// TIA Portal project "State Machine Triple-liquid mixing+HMI final version" (V17)

(* hardware
DEVICE "S7-300/ET200M station_1"  S7-300 station
   slot 0: "Rail_0"  Rail  6ES7 390-1***0-0AA0
   slot 2: "PLC_1"  CPU 317-2 PN/DP  6ES7 317-2EK14-0AB0  V3.2
      slot 2: "PROFINET interface_1"  PN-IO
         slot 1: "Port_1"  Port
         slot 2: "Port_2"  Port
   slot 4: "DI 16x24VDC_1"  DI16 x 24VDC  6ES7 321-1BH02-0AA0
   slot 5: "DO 8x24VDC/0.5A_1"  DO8 x 24VDC / 0.5A  6ES7 322-8BF00-0AB0
   slot 6: "AI 4x0/4mA/20mA, Ex_1"  AI4 x 0/4 to 20mA, Ex  6ES7 331-7RD00-0AB0
DEVICE "HMI_1"  TP1200 Comfort Portrait SIPLUS
   slot 0: "HMI_1"  TP1200 Comfort Portrait SIPLUS  6AG1 124-0MC01-4AX0  17.0.0.0
   slot 1: "HMI_RT_1"  TP1200 Comfort Portrait SIPLUS  6AG1 124-0MC01-4AX0  17.0.0.0
   slot 5: "HMI_1.IE_CP_1"  PROFINET Interface  17.0.0.0
      slot 1: "PROFINET Interface_1"  PROFINET Interface
         slot 1: "Port_1"  Port
         slot 2: "Port_2"  Port
   slot 7: "HMI_1.MPI/DP_CP_1"  MPI/DP Interface  17.0.0.0
*)

// ===== PLC "PLC_1"  CPU 317-2 PN/DP =====

VAR_GLOBAL   // PLC tag table "Default tag table"
   "E_stop" AT %I0.0 : Bool;
   "Actual_level" AT %MD0 : Real;
   "RESET_1" AT %I0.1 : Bool;
   "Start_mixing" AT %I0.2 : Bool;
   "Alarm_light" AT %Q0.0 : Bool;
   "Valve_A" AT %Q4.0 : Bool;
   "Valve_B" AT %Q4.1 : Bool;
   "Valve_C" AT %Q4.2 : Bool;
   "Agitator_Q" AT %Q4.3 : Bool;
   "Drain_valve" AT %Q4.4 : Bool;
   "REC_A" AT %MD4 : Real;
   "REC_B" AT %MD8 : Real;
   "REC_C" AT %MD12 : Real;
   "start_empty" AT %I0.3 : Bool;
   "Eroor_code" AT %MW16 : Int;
   "Start_timer" AT %T0 : Timer;
   "start_empty_Timer" AT %T1 : Timer;
   "Reset_timer" AT %T2 : Timer;
   "RAW_Level_sensor" AT %IW288 : Int;
   "Start_batch" AT %M10.1 : Bool;
   "Reset_HMI" AT %M10.2 : Bool;
   "Start-EMpty" AT %M10.3 : Bool;
   "Status" AT %MW20 : Int;
   "Min_level" AT %MD48 : Real;
   "Max_lvl" AT %MD24 : Real;
   "drain_time_WD" AT %MD28 : Time;
   "Agitator_time_WD" AT %MD32 : Time;
   "FIlling_time_WD" AT %MD36 : Time;
   "Agitating_time" AT %MD40 : Time;
   "Batch_done_confirmation" AT %M44.0 : Bool;
   "Rec_approved" AT %M44.1 : Bool;
   "Tank1_active" AT %M18.0 : Bool;
   "Alarm_HMI" AT %M18.1 : Bool;
   "Valv_A_HMI" AT %M18.2 : Bool;
   "Valv_B_HMI" AT %M18.3 : Bool;
   "Valv_C_HMI" AT %M18.4 : Bool;
   "Agit_HMI" AT %M18.5 : Bool;
   "Drain_valv_HMI" AT %M18.6 : Bool;
END_VAR

DATA_BLOCK "batch_variable"   // DB9
{ S7_Optimized_Access := 'FALSE' }
VERSION : 0.1
   VAR
      reciepe_A : Real;
      reciepe_B : Real;
      reciepe_C : Real;
   END_VAR
BEGIN
END_DATA_BLOCK

DATA_BLOCK "Stat machine_DB"   // DB10
{ S7_Optimized_Access := 'FALSE' }
VERSION : 0.1
// stored: InstanceOfName Stat machine
"Stat machine"
BEGIN
END_DATA_BLOCK

FUNCTION_BLOCK "Stat machine"   // FB1, LAD
{ S7_Optimized_Access := 'FALSE' }
VERSION : 0.1
   VAR_INPUT
      "E-Stop" : Bool;
      Actual_level : Real;
      RESET_Cmd : Bool;
      start_mixing : Bool;
      Reciepes_A : Real;
      Reciepes_c : Real;
      Reciepes_B : Real;
      start_empty : Bool;
      wtachDog_time_Drain : Time;
      wtachDog_time_Agitator : Time;
      wtachDog_time_valve : Time;
      Min_level : Real;
      Agitating_time : Time;
      batch_done_confirmation : Bool;
   END_VAR
   VAR_OUTPUT
      Alram_red_light : Bool;
      q_valve_A : Bool;
      q_valve_B : Bool;
      q_valve_C : Bool;
      Agitaor : Bool;
      drain_valve : Bool;
      Error_code : Int;
      Alarm_active : Bool;
      Valve_A_active : Bool;
      Valve_B_active : Bool;
      Valve_C_active : Bool;
      Agitator_active : Bool;
      Drain_valve_active : Bool;
   END_VAR
   VAR_IN_OUT
      iStep_number : Int;
      max_lvl : Real;
      Recrp_approved : Bool;
   END_VAR
   VAR
      Agitator_runnig : Bool;
      Target_1 : Real;
      Target_2 : Real;
      Reset_alrm : Bool;
      Batch_done : Bool;
      "1%_tank_apacity" : Real;
      max_recepes_valuem : Real;
      "15%_Tank_capacity" : Real;
   END_VAR
   VAR_TEMP   // added for the SCL form of the ladder/FBD networks
      _w1 : Bool;
   END_VAR
BEGIN

REGION Network 1
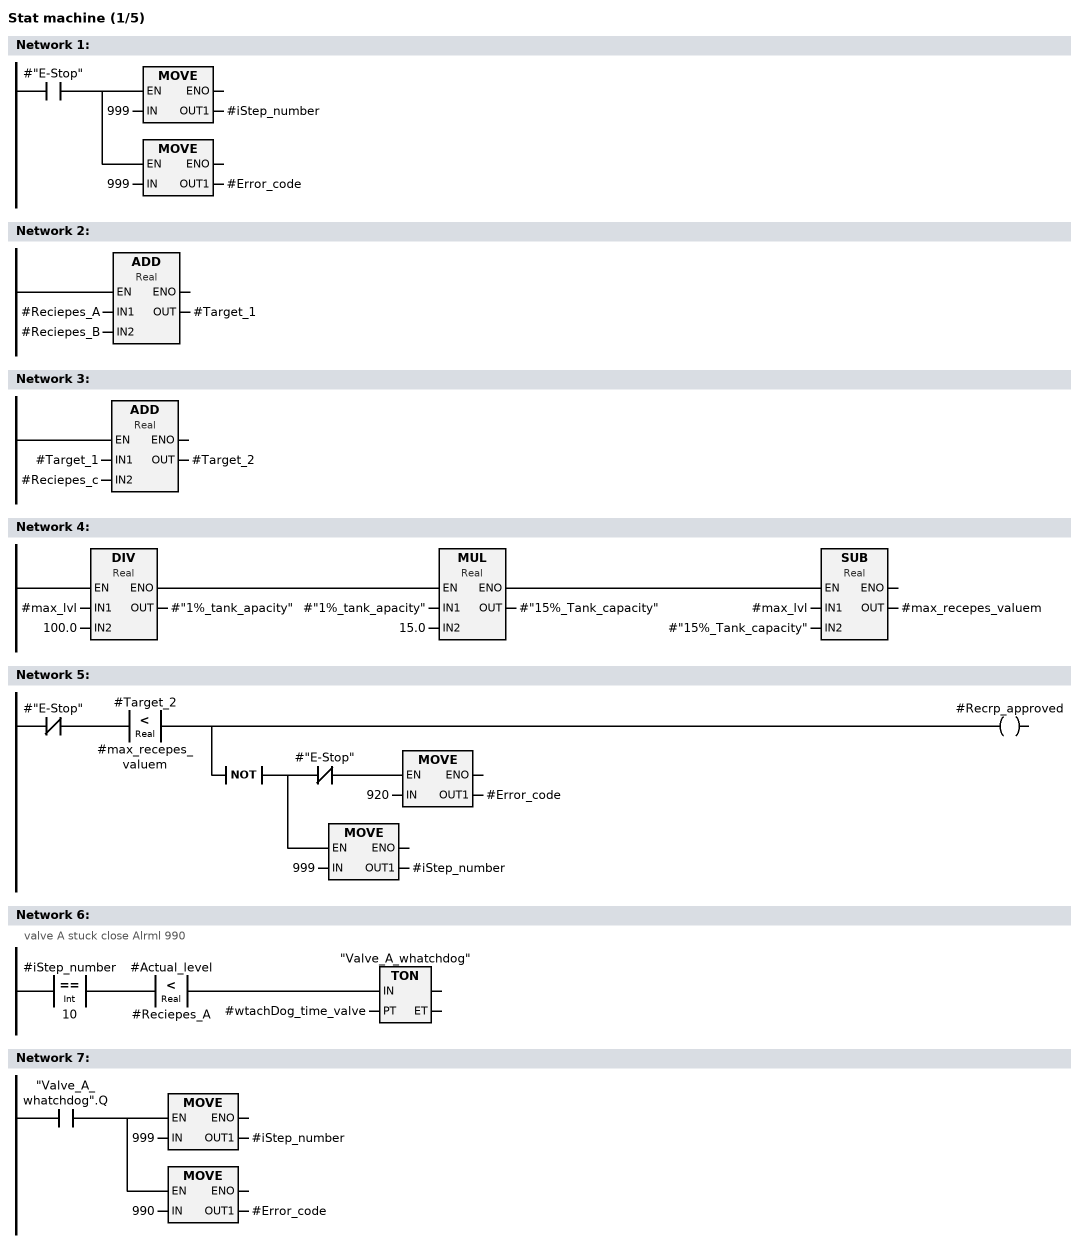
   RUNG wire#powerrail
      Contact( #"E-Stop" )
      wire#w1
      { S7_GenerateENO := "TRUE" } Move(in := 999, out1 => #iStep_number)
   END_RUNG
   RUNG wire#w1
      { S7_GenerateENO := "TRUE" } Move(in := 999, out1 => #Error_code)
   END_RUNG
   // the same network as SCL:
   IF #"E-Stop" THEN
       #iStep_number := 999;
       #Error_code := 999;
   END_IF;
END_REGION

REGION Network 2
   RUNG wire#powerrail
      { S7_Templates := "SrcType := Real"; S7_GenerateENO := "TRUE" } Add(in1 := #Reciepes_A, in2 := #Reciepes_B, out => #Target_1)
   END_RUNG
   // the same network as SCL:
   #Target_1 := #Reciepes_A + #Reciepes_B;
END_REGION

REGION Network 3
   RUNG wire#powerrail
      { S7_Templates := "SrcType := Real"; S7_GenerateENO := "TRUE" } Add(in1 := #Target_1, in2 := #Reciepes_c, out => #Target_2)
   END_RUNG
   // the same network as SCL:
   #Target_2 := #Target_1 + #Reciepes_c;
END_REGION

REGION Network 4
   RUNG wire#powerrail
      { S7_Templates := "SrcType := Real"; S7_GenerateENO := "TRUE" } Div(in1 := #max_lvl, in2 := 100.0, out => #"1%_tank_apacity")
      { S7_Templates := "SrcType := Real"; S7_GenerateENO := "TRUE" } Mul(in1 := #"1%_tank_apacity", in2 := 15.0, out => #"15%_Tank_capacity")
      { S7_Templates := "SrcType := Real"; S7_GenerateENO := "TRUE" } Sub(in1 := #max_lvl, in2 := #"15%_Tank_capacity", out => #max_recepes_valuem)
   END_RUNG
   // the same network as SCL:
   // ENO of a box is taken as its EN; it also drops when the box reports an error
   #"1%_tank_apacity" := #max_lvl / 100.0;
   #"15%_Tank_capacity" := #"1%_tank_apacity" * 15.0;
   #max_recepes_valuem := #max_lvl - #"15%_Tank_capacity";
END_REGION

REGION Network 5
   RUNG wire#powerrail
      I_Contact( #"E-Stop" )
      { S7_Templates := "SrcType := Real" } LT_Contact(in1 := #Target_2, in2 := #max_recepes_valuem)
      wire#w1
      Coil( #Recrp_approved )
   END_RUNG
   RUNG wire#w1
      Not()
      wire#w2
      I_Contact( #"E-Stop" )
      { S7_GenerateENO := "TRUE" } Move(in := 920, out1 => #Error_code)
   END_RUNG
   RUNG wire#w2
      { S7_GenerateENO := "TRUE" } Move(in := 999, out1 => #iStep_number)
   END_RUNG
   // the same network as SCL:
   #Recrp_approved := NOT #"E-Stop" AND (#Target_2 < #max_recepes_valuem);
   IF NOT #Recrp_approved AND NOT #"E-Stop" THEN #Error_code := 920; END_IF;
   IF NOT #Recrp_approved THEN #iStep_number := 999; END_IF;
END_REGION

REGION Network 6
   // valve A stuck close Alrml 990
   "Valve_A_whatchdog".TON(IN := (#iStep_number = 10) AND (#Actual_level < #Reciepes_A),
                           PT := #wtachDog_time_valve);
END_REGION

REGION Network 7
   RUNG wire#powerrail
      Contact( "Valve_A_whatchdog".Q )
      wire#w1
      { S7_GenerateENO := "TRUE" } Move(in := 999, out1 => #iStep_number)
   END_RUNG
   RUNG wire#w1
      { S7_GenerateENO := "TRUE" } Move(in := 990, out1 => #Error_code)
   END_RUNG
   // the same network as SCL:
   IF "Valve_A_whatchdog".Q THEN
       #iStep_number := 999;
       #Error_code := 990;
   END_IF;
END_REGION

REGION Network 8
   // valve B stuck open alrm 989
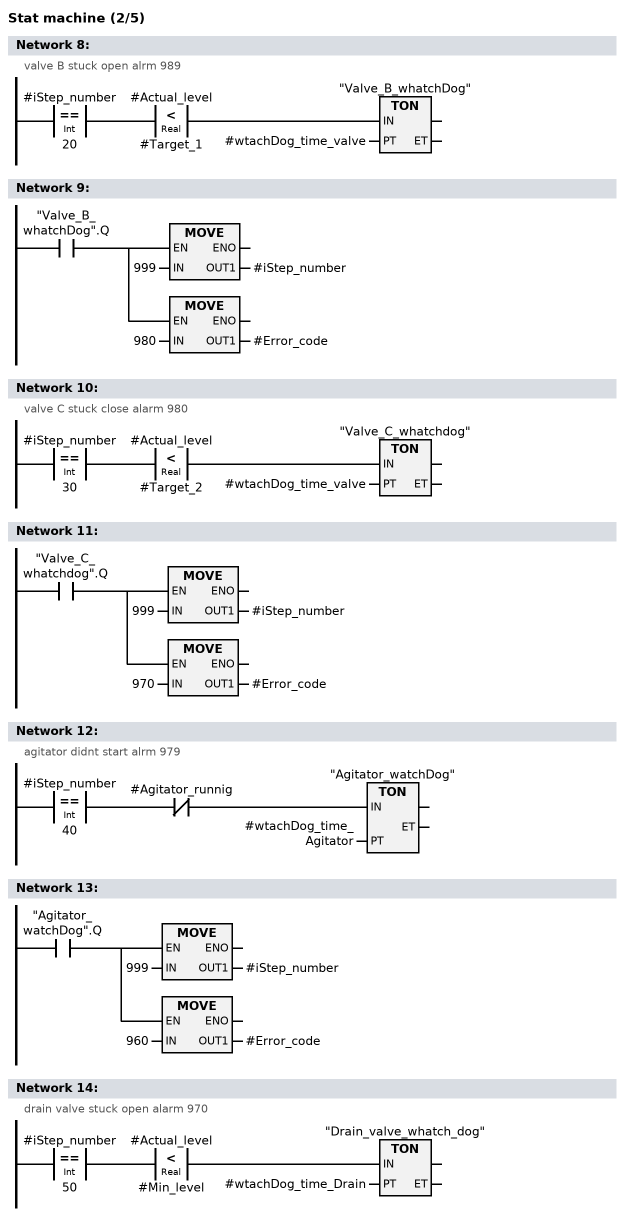
   "Valve_B_whatchDog".TON(IN := (#iStep_number = 20) AND (#Actual_level < #Target_1),
                           PT := #wtachDog_time_valve);
END_REGION

REGION Network 9
   RUNG wire#powerrail
      Contact( "Valve_B_whatchDog".Q )
      wire#w1
      { S7_GenerateENO := "TRUE" } Move(in := 999, out1 => #iStep_number)
   END_RUNG
   RUNG wire#w1
      { S7_GenerateENO := "TRUE" } Move(in := 980, out1 => #Error_code)
   END_RUNG
   // the same network as SCL:
   IF "Valve_B_whatchDog".Q THEN
       #iStep_number := 999;
       #Error_code := 980;
   END_IF;
END_REGION

REGION Network 10
   // valve C stuck close alarm 980
   "Valve_C_whatchdog".TON(IN := (#iStep_number = 30) AND (#Actual_level < #Target_2),
                           PT := #wtachDog_time_valve);
END_REGION

REGION Network 11
   RUNG wire#powerrail
      Contact( "Valve_C_whatchdog".Q )
      wire#w1
      { S7_GenerateENO := "TRUE" } Move(in := 999, out1 => #iStep_number)
   END_RUNG
   RUNG wire#w1
      { S7_GenerateENO := "TRUE" } Move(in := 970, out1 => #Error_code)
   END_RUNG
   // the same network as SCL:
   IF "Valve_C_whatchdog".Q THEN
       #iStep_number := 999;
       #Error_code := 970;
   END_IF;
END_REGION

REGION Network 12
   // agitator didnt start alrm 979
   "Agitator_watchDog".TON(IN := (#iStep_number = 40) AND NOT #Agitator_runnig, PT := #wtachDog_time_Agitator);
END_REGION

REGION Network 13
   RUNG wire#powerrail
      Contact( "Agitator_watchDog".Q )
      wire#w1
      { S7_GenerateENO := "TRUE" } Move(in := 999, out1 => #iStep_number)
   END_RUNG
   RUNG wire#w1
      { S7_GenerateENO := "TRUE" } Move(in := 960, out1 => #Error_code)
   END_RUNG
   // the same network as SCL:
   IF "Agitator_watchDog".Q THEN
       #iStep_number := 999;
       #Error_code := 960;
   END_IF;
END_REGION

REGION Network 14
   // drain valve stuck open alarm 970
   "Drain_valve_whatch_dog".TON(IN := (#iStep_number = 50) AND (#Actual_level < #Min_level),
                           PT := #wtachDog_time_Drain);
END_REGION

REGION Network 15
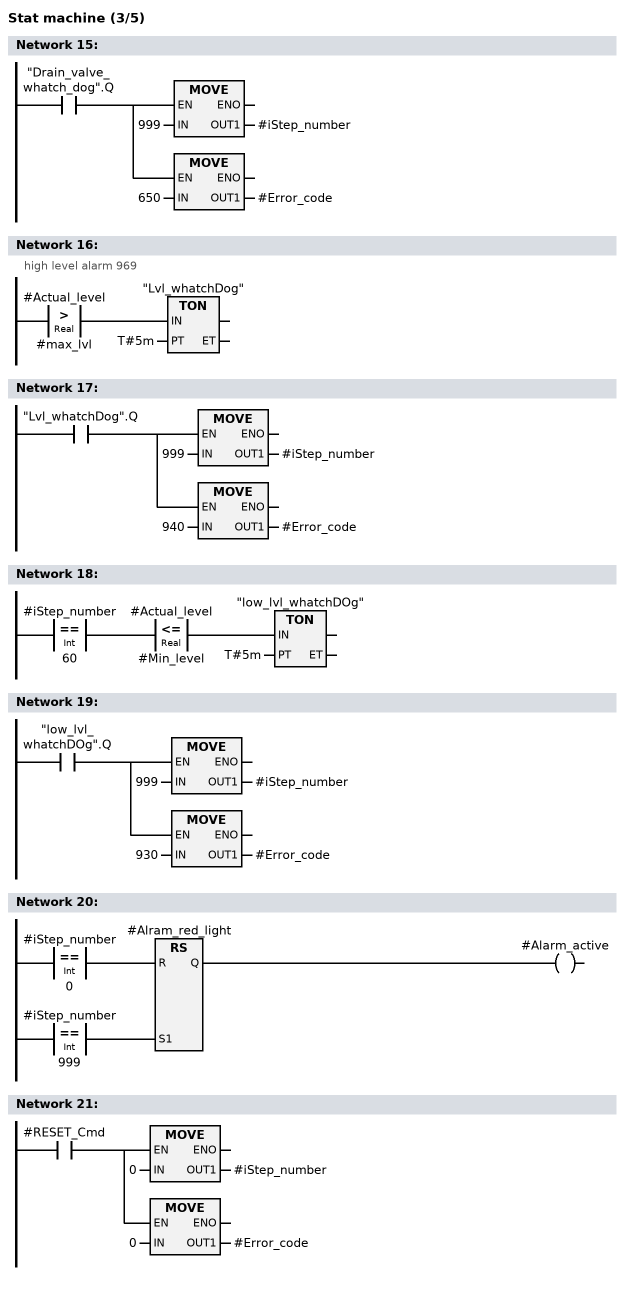
   RUNG wire#powerrail
      Contact( "Drain_valve_whatch_dog".Q )
      wire#w1
      { S7_GenerateENO := "TRUE" } Move(in := 999, out1 => #iStep_number)
   END_RUNG
   RUNG wire#w1
      { S7_GenerateENO := "TRUE" } Move(in := 650, out1 => #Error_code)
   END_RUNG
   // the same network as SCL:
   IF "Drain_valve_whatch_dog".Q THEN
       #iStep_number := 999;
       #Error_code := 650;
   END_IF;
END_REGION

REGION Network 16
   // high level alarm 969
   "Lvl_whatchDog".TON(IN := #Actual_level > #max_lvl, PT := T#5m);
END_REGION

REGION Network 17
   RUNG wire#powerrail
      Contact( "Lvl_whatchDog".Q )
      wire#w1
      { S7_GenerateENO := "TRUE" } Move(in := 999, out1 => #iStep_number)
   END_RUNG
   RUNG wire#w1
      { S7_GenerateENO := "TRUE" } Move(in := 940, out1 => #Error_code)
   END_RUNG
   // the same network as SCL:
   IF "Lvl_whatchDog".Q THEN
       #iStep_number := 999;
       #Error_code := 940;
   END_IF;
END_REGION

REGION Network 18
   "low_lvl_whatchDOg".TON(IN := (#iStep_number = 60) AND (#Actual_level <= #Min_level), PT := T#5m);
END_REGION

REGION Network 19
   RUNG wire#powerrail
      Contact( "low_lvl_whatchDOg".Q )
      wire#w1
      { S7_GenerateENO := "TRUE" } Move(in := 999, out1 => #iStep_number)
   END_RUNG
   RUNG wire#w1
      { S7_GenerateENO := "TRUE" } Move(in := 930, out1 => #Error_code)
   END_RUNG
   // the same network as SCL:
   IF "low_lvl_whatchDOg".Q THEN
       #iStep_number := 999;
       #Error_code := 930;
   END_IF;
END_REGION

REGION Network 20
   RUNG wire#powerrail
      { S7_Templates := "SrcType := Int" } EQ_Contact(in1 := #iStep_number, in2 := 0)
      S_RS(operand := #Alram_red_light, s1 := wire#w1)
      Coil( #Alarm_active )
   END_RUNG
   RUNG wire#powerrail
      { S7_Templates := "SrcType := Int" } EQ_Contact(in1 := #iStep_number, in2 := 999)
   END_RUNG wire#w1
   // the same network as SCL:
   IF #iStep_number = 0 THEN
       #Alram_red_light := FALSE;   // RS flip-flop
   END_IF;
   IF #iStep_number = 999 THEN #Alram_red_light := TRUE; END_IF;
   #Alarm_active := #Alram_red_light;
END_REGION

REGION Network 21
   RUNG wire#powerrail
      Contact( #RESET_Cmd )
      wire#w1
      { S7_GenerateENO := "TRUE" } Move(in := 0, out1 => #iStep_number)
   END_RUNG
   RUNG wire#w1
      { S7_GenerateENO := "TRUE" } Move(in := 0, out1 => #Error_code)
   END_RUNG
   // the same network as SCL:
   IF #RESET_Cmd THEN
       #iStep_number := 0;
       #Error_code := 0;
   END_IF;
END_REGION

REGION Network 22
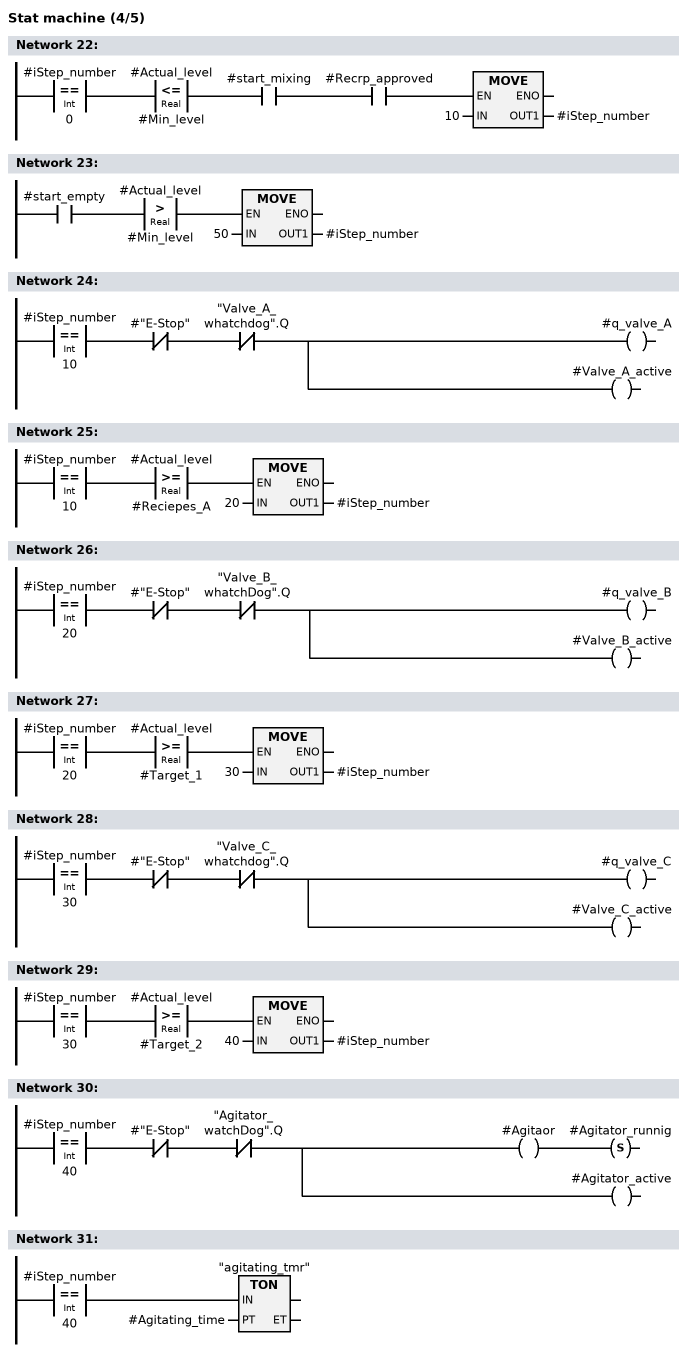
   RUNG wire#powerrail
      { S7_Templates := "SrcType := Int" } EQ_Contact(in1 := #iStep_number, in2 := 0)
      { S7_Templates := "SrcType := Real" } LE_Contact(in1 := #Actual_level, in2 := #Min_level)
      Contact( #start_mixing )
      Contact( #Recrp_approved )
      { S7_GenerateENO := "TRUE" } Move(in := 10, out1 => #iStep_number)
   END_RUNG
   // the same network as SCL:
   IF (#iStep_number = 0) AND (#Actual_level <= #Min_level) AND #start_mixing AND #Recrp_approved THEN
       #iStep_number := 10;
   END_IF;
END_REGION

REGION Network 23
   RUNG wire#powerrail
      Contact( #start_empty )
      { S7_Templates := "SrcType := Real" } GT_Contact(in1 := #Actual_level, in2 := #Min_level)
      { S7_GenerateENO := "TRUE" } Move(in := 50, out1 => #iStep_number)
   END_RUNG
   // the same network as SCL:
   IF #start_empty AND (#Actual_level > #Min_level) THEN #iStep_number := 50; END_IF;
END_REGION

REGION Network 24
   RUNG wire#powerrail
      { S7_Templates := "SrcType := Int" } EQ_Contact(in1 := #iStep_number, in2 := 10)
      I_Contact( #"E-Stop" )
      I_Contact( "Valve_A_whatchdog".Q )
      wire#w1
      Coil( #q_valve_A )
   END_RUNG
   RUNG wire#w1
      Coil( #Valve_A_active )
   END_RUNG
   // the same network as SCL:
   #q_valve_A := (#iStep_number = 10) AND NOT #"E-Stop" AND NOT "Valve_A_whatchdog".Q;
   #Valve_A_active := #q_valve_A;
END_REGION

REGION Network 25
   RUNG wire#powerrail
      { S7_Templates := "SrcType := Int" } EQ_Contact(in1 := #iStep_number, in2 := 10)
      { S7_Templates := "SrcType := Real" } GE_Contact(in1 := #Actual_level, in2 := #Reciepes_A)
      { S7_GenerateENO := "TRUE" } Move(in := 20, out1 => #iStep_number)
   END_RUNG
   // the same network as SCL:
   IF (#iStep_number = 10) AND (#Actual_level >= #Reciepes_A) THEN #iStep_number := 20; END_IF;
END_REGION

REGION Network 26
   RUNG wire#powerrail
      { S7_Templates := "SrcType := Int" } EQ_Contact(in1 := #iStep_number, in2 := 20)
      I_Contact( #"E-Stop" )
      I_Contact( "Valve_B_whatchDog".Q )
      wire#w1
      Coil( #q_valve_B )
   END_RUNG
   RUNG wire#w1
      Coil( #Valve_B_active )
   END_RUNG
   // the same network as SCL:
   #q_valve_B := (#iStep_number = 20) AND NOT #"E-Stop" AND NOT "Valve_B_whatchDog".Q;
   #Valve_B_active := #q_valve_B;
END_REGION

REGION Network 27
   RUNG wire#powerrail
      { S7_Templates := "SrcType := Int" } EQ_Contact(in1 := #iStep_number, in2 := 20)
      { S7_Templates := "SrcType := Real" } GE_Contact(in1 := #Actual_level, in2 := #Target_1)
      { S7_GenerateENO := "TRUE" } Move(in := 30, out1 => #iStep_number)
   END_RUNG
   // the same network as SCL:
   IF (#iStep_number = 20) AND (#Actual_level >= #Target_1) THEN #iStep_number := 30; END_IF;
END_REGION

REGION Network 28
   RUNG wire#powerrail
      { S7_Templates := "SrcType := Int" } EQ_Contact(in1 := #iStep_number, in2 := 30)
      I_Contact( #"E-Stop" )
      I_Contact( "Valve_C_whatchdog".Q )
      wire#w1
      Coil( #q_valve_C )
   END_RUNG
   RUNG wire#w1
      Coil( #Valve_C_active )
   END_RUNG
   // the same network as SCL:
   #q_valve_C := (#iStep_number = 30) AND NOT #"E-Stop" AND NOT "Valve_C_whatchdog".Q;
   #Valve_C_active := #q_valve_C;
END_REGION

REGION Network 29
   RUNG wire#powerrail
      { S7_Templates := "SrcType := Int" } EQ_Contact(in1 := #iStep_number, in2 := 30)
      { S7_Templates := "SrcType := Real" } GE_Contact(in1 := #Actual_level, in2 := #Target_2)
      { S7_GenerateENO := "TRUE" } Move(in := 40, out1 => #iStep_number)
   END_RUNG
   // the same network as SCL:
   IF (#iStep_number = 30) AND (#Actual_level >= #Target_2) THEN #iStep_number := 40; END_IF;
END_REGION

REGION Network 30
   RUNG wire#powerrail
      { S7_Templates := "SrcType := Int" } EQ_Contact(in1 := #iStep_number, in2 := 40)
      I_Contact( #"E-Stop" )
      I_Contact( "Agitator_watchDog".Q )
      wire#w1
      Coil( #Agitaor )
      S_Coil( #Agitator_runnig )
   END_RUNG
   RUNG wire#w1
      Coil( #Agitator_active )
   END_RUNG
   // the same network as SCL:
   #Agitaor := (#iStep_number = 40) AND NOT #"E-Stop" AND NOT "Agitator_watchDog".Q;
   IF #Agitaor THEN #Agitator_runnig := TRUE; END_IF;
   #Agitator_active := #Agitaor;
END_REGION

REGION Network 31
   "agitating_tmr".TON(IN := #iStep_number = 40, PT := #Agitating_time);
END_REGION

REGION Network 32
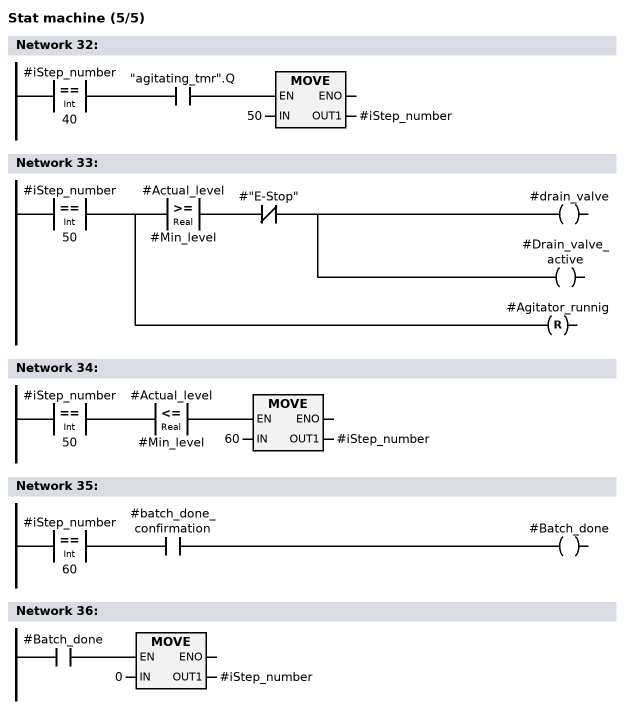
   RUNG wire#powerrail
      { S7_Templates := "SrcType := Int" } EQ_Contact(in1 := #iStep_number, in2 := 40)
      Contact( "agitating_tmr".Q )
      { S7_GenerateENO := "TRUE" } Move(in := 50, out1 => #iStep_number)
   END_RUNG
   // the same network as SCL:
   IF (#iStep_number = 40) AND "agitating_tmr".Q THEN #iStep_number := 50; END_IF;
END_REGION

REGION Network 33
   RUNG wire#powerrail
      { S7_Templates := "SrcType := Int" } EQ_Contact(in1 := #iStep_number, in2 := 50)
      wire#w1
      { S7_Templates := "SrcType := Real" } GE_Contact(in1 := #Actual_level, in2 := #Min_level)
      I_Contact( #"E-Stop" )
      wire#w2
      Coil( #drain_valve )
   END_RUNG
   RUNG wire#w2
      Coil( #Drain_valve_active )
   END_RUNG
   RUNG wire#w1
      R_Coil( #Agitator_runnig )
   END_RUNG
   // the same network as SCL:
   #_w1 := #iStep_number = 50;
   #drain_valve := #_w1 AND (#Actual_level >= #Min_level) AND NOT #"E-Stop";
   #Drain_valve_active := #drain_valve;
   IF #_w1 THEN #Agitator_runnig := FALSE; END_IF;
END_REGION

REGION Network 34
   RUNG wire#powerrail
      { S7_Templates := "SrcType := Int" } EQ_Contact(in1 := #iStep_number, in2 := 50)
      { S7_Templates := "SrcType := Real" } LE_Contact(in1 := #Actual_level, in2 := #Min_level)
      { S7_GenerateENO := "TRUE" } Move(in := 60, out1 => #iStep_number)
   END_RUNG
   // the same network as SCL:
   IF (#iStep_number = 50) AND (#Actual_level <= #Min_level) THEN #iStep_number := 60; END_IF;
END_REGION

REGION Network 35
   RUNG wire#powerrail
      { S7_Templates := "SrcType := Int" } EQ_Contact(in1 := #iStep_number, in2 := 60)
      Contact( #batch_done_confirmation )
      Coil( #Batch_done )
   END_RUNG
   // the same network as SCL:
   #Batch_done := (#iStep_number = 60) AND #batch_done_confirmation;
END_REGION

REGION Network 36
   RUNG wire#powerrail
      Contact( #Batch_done )
      { S7_GenerateENO := "TRUE" } Move(in := 0, out1 => #iStep_number)
   END_RUNG
   // the same network as SCL:
   IF #Batch_done THEN #iStep_number := 0; END_IF;
END_REGION
END_FUNCTION_BLOCK

FUNCTION "Level_sensor" : Void   // FC1, LAD
{ S7_Optimized_Access := 'FALSE' }
VERSION : 0.1
   VAR_INPUT
      Raw_sensro : Int;
   END_VAR
   VAR_OUTPUT
      Scaled_value : Real;
   END_VAR
   VAR_TEMP
      false_1 : Bool;
      Error_1 : Word;
   END_VAR
BEGIN

REGION Network 1
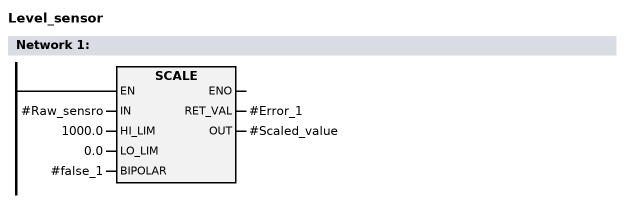
   #Error_1 := SCALE(IN := #Raw_sensro,
                     HI_LIM := 1000.0,
                     LO_LIM := 0.0,
                     BIPOLAR := #false_1,
                     OUT => #Scaled_value);
END_REGION
END_FUNCTION

ORGANIZATION_BLOCK "Main"   // OB1, LAD
TITLE = "Main Program Sweep (Cycle)"
{ S7_Optimized_Access := 'FALSE' }
VERSION : 0.1
   VAR_TEMP
      OB1_EV_CLASS : Byte;   // Bits 0-3 = 1 (Coming event), Bits 4-7 = 1 (Event class 1)
      OB1_SCAN_1 : Byte;   // 1 (Cold restart scan 1 of OB 1), 3 (Scan 2-n of OB 1)
      OB1_PRIORITY : Byte;   // Priority of OB Execution
      OB1_OB_NUMBR : Byte;   // 1 (Organization block 1, OB1)
      OB1_RESERVED_1 : Byte;   // Reserved for system
      OB1_RESERVED_2 : Byte;   // Reserved for system
      OB1_PREV_CYCLE : Int;   // Cycle time of previous OB1 scan (milliseconds)
      OB1_MIN_CYCLE : Int;   // Minimum cycle time of OB1 (milliseconds)
      OB1_MAX_CYCLE : Int;   // Maximum cycle time of OB1 (milliseconds)
      OB1_DATE_TIME : Date_And_Time;   // Date and time OB1 started
   END_VAR
   VAR_TEMP   // added for the SCL form of the ladder/FBD networks
      _w1 : Bool;
      _s5time1 : S5Time;
      _w2 : Bool;
      _s5time2 : S5Time;
      _w3 : Bool;
      _s5time3 : S5Time;
      _w4 : Bool;
   END_VAR
BEGIN

REGION Network 1
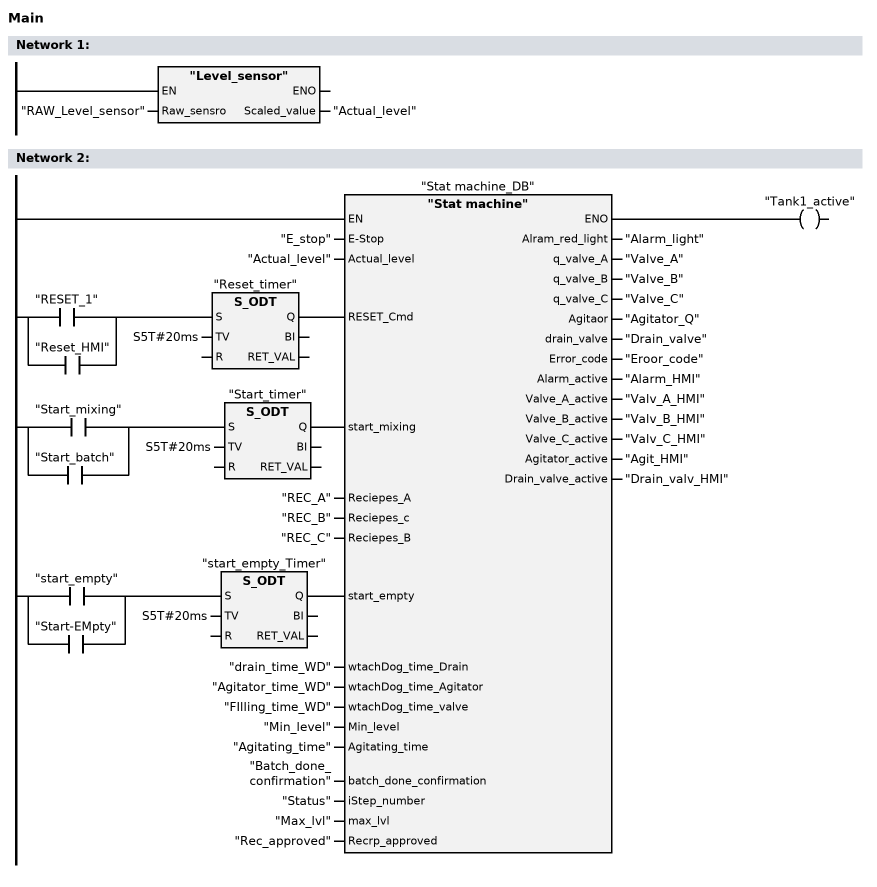
   RUNG wire#powerrail
      "Level_sensor"(Raw_sensro := "RAW_Level_sensor", Scaled_value => "Actual_level")
   END_RUNG
   // the same network as SCL:
   "Level_sensor"(Raw_sensro := "RAW_Level_sensor", Scaled_value => "Actual_level");
END_REGION

REGION Network 2
   RUNG wire#powerrail
      "Stat machine_DB"(RESET_Cmd := wire#w2, start_mixing := wire#w4, start_empty := wire#w6, "E-Stop" := "E_stop", Actual_level := "Actual_level", Reciepes_A := "REC_A", Reciepes_c := "REC_B", Reciepes_B := "REC_C", wtachDog_time_Drain := "drain_time_WD", wtachDog_time_Agitator := "Agitator_time_WD", wtachDog_time_valve := "FIlling_time_WD", Min_level := "Min_level", Agitating_time := "Agitating_time", batch_done_confirmation := "Batch_done_confirmation", iStep_number := "Status", max_lvl := "Max_lvl", Recrp_approved := "Rec_approved", Alram_red_light => "Alarm_light", q_valve_A => "Valve_A", q_valve_B => "Valve_B", q_valve_C => "Valve_C", Agitaor => "Agitator_Q", drain_valve => "Drain_valve", Error_code => "Eroor_code", Alarm_active => "Alarm_HMI", Valve_A_active => "Valv_A_HMI", Valve_B_active => "Valv_B_HMI", Valve_C_active => "Valv_C_HMI", Agitator_active => "Agit_HMI", Drain_valve_active => "Drain_valv_HMI")
      Coil( "Tank1_active" )
   END_RUNG
   RUNG wire#powerrail
      Contact( "RESET_1" )
      wire#w1
      S_ODT(T_NO := "Reset_timer", TV := S5T#20ms, R :=, BI =>, RET_VAL =>)
   END_RUNG wire#w2
   RUNG wire#powerrail
      Contact( "Reset_HMI" )
   END_RUNG wire#w1
   RUNG wire#powerrail
      Contact( "Start_mixing" )
      wire#w3
      S_ODT(T_NO := "Start_timer", TV := S5T#20ms, R :=, BI =>, RET_VAL =>)
   END_RUNG wire#w4
   RUNG wire#powerrail
      Contact( "Start_batch" )
   END_RUNG wire#w3
   RUNG wire#powerrail
      Contact( "start_empty" )
      wire#w5
      S_ODT(T_NO := "start_empty_Timer", TV := S5T#20ms, R :=, BI =>, RET_VAL =>)
   END_RUNG wire#w6
   RUNG wire#powerrail
      Contact( "Start-EMpty" )
   END_RUNG wire#w5
   // the same network as SCL:
   #_s5time1 := S_ODT(T_NO := "Reset_timer", S := "RESET_1" OR "Reset_HMI", TV := S5T#20ms, Q => #_w1);
   #_s5time2 := S_ODT(T_NO := "Start_timer", S := "Start_mixing" OR "Start_batch", TV := S5T#20ms, Q => #_w2);
   #_s5time3 := S_ODT(T_NO := "start_empty_Timer",
                      S := "start_empty" OR "Start-EMpty",
                      TV := S5T#20ms,
                      Q => #_w3);
   "Stat machine_DB"("E-Stop" := "E_stop",   // "Stat machine"
                     Actual_level := "Actual_level",
                     RESET_Cmd := #_w1,
                     start_mixing := #_w2,
                     Reciepes_A := "REC_A",
                     Reciepes_c := "REC_B",
                     Reciepes_B := "REC_C",
                     start_empty := #_w3,
                     wtachDog_time_Drain := "drain_time_WD",
                     wtachDog_time_Agitator := "Agitator_time_WD",
                     wtachDog_time_valve := "FIlling_time_WD",
                     Min_level := "Min_level",
                     Agitating_time := "Agitating_time",
                     batch_done_confirmation := "Batch_done_confirmation",
                     iStep_number := "Status",
                     max_lvl := "Max_lvl",
                     Recrp_approved := "Rec_approved",
                     Alram_red_light => "Alarm_light",
                     q_valve_A => "Valve_A",
                     q_valve_B => "Valve_B",
                     q_valve_C => "Valve_C",
                     Agitaor => "Agitator_Q",
                     drain_valve => "Drain_valve",
                     Error_code => "Eroor_code",
                     Alarm_active => "Alarm_HMI",
                     Valve_A_active => "Valv_A_HMI",
                     Valve_B_active => "Valv_B_HMI",
                     Valve_C_active => "Valv_C_HMI",
                     Agitator_active => "Agit_HMI",
                     Drain_valve_active => "Drain_valv_HMI",
                     ENO => #_w4);
   "Tank1_active" := #_w4;
END_REGION
END_ORGANIZATION_BLOCK

ORGANIZATION_BLOCK "COMPLETE RESTART"   // OB100, LAD
TITLE = "Complete Restart"
{ S7_Optimized_Access := 'FALSE' }
VERSION : 0.1
   VAR_TEMP
      OB100_EV_CLASS : Byte;   // 16#13, Event class 1, Entering event state, Event logged in diagnostic buffer
      OB100_STRTUP : Byte;   // 16#81/82/83/84 Method of startup
      OB100_PRIORITY : Byte;   // Priority of OB Execution
      OB100_OB_NUMBR : Byte;   // 100 (Organization block 100, OB100)
      OB100_RESERVED_1 : Byte;   // Reserved for system
      OB100_RESERVED_2 : Byte;   // Reserved for system
      OB100_STOP : Word;   // Event that caused CPU to stop (16#4xxx)
      OB100_STRT_INFO : DWord;   // Information on how system started
      OB100_DATE_TIME : Date_And_Time;   // Date and time OB100 started
   END_VAR
BEGIN

REGION Network 1
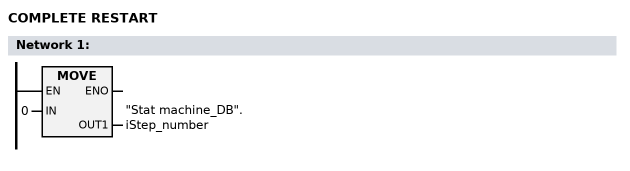
   RUNG wire#powerrail
      { S7_GenerateENO := "TRUE" } Move(in := 0, out1 => "Stat machine_DB".iStep_number)
   END_RUNG
   // the same network as SCL:
   "Stat machine_DB".iStep_number := 0;
END_REGION
END_ORGANIZATION_BLOCK

(* ===== HMI "HMI_RT_1" =====
system functions are stored by id; their names below are inferred from use
connection "Connection_1": ETHERNET, SIMATIC S7 300/400 MPI
connection "HMI_Connection_1": ETHERNET, SIMATIC S7 300/400 MPI

HMI tags "Default tag table"
   "Start_Batch" : Bool = PLC Start_batch AT %M10.1, 1 s
   "Reset_HMI" : Bool = PLC Reset_HMI AT %M10.2, 1 s
   "Star_empty" : Bool = PLC "Start-EMpty" AT %M10.3, 1 s
   "level_value" : Real = PLC Actual_level AT %MD0, 1 s
   "Error_code" : Int = PLC Eroor_code AT %MW16, 1 s
   "Recipes_A" : Real = PLC REC_A AT %MD4, 1 s
   "Recipes_B" : Real = PLC REC_B AT %MD8, 1 s
   "Recipes_C" : Real = PLC REC_C AT %MD12, 1 s
   "Status" : Int = PLC Status AT %MW20, 1 s
   "max _lvl" : Real = PLC Max_lvl AT %MD24, 1 s
   "min_lvl" : Real = PLC Min_level AT %MD48, 1 s
   "drain_time_WD" : Time = PLC drain_time_WD AT %MD28, 1 s
   "Agitator_time_WD" : Time = PLC Agitator_time_WD AT %MD32, 1 s
   "agitating_time" : Time = PLC Agitating_time AT %MD40, 1 s
   "filling_time_WD" : Time = PLC FIlling_time_WD AT %MD36, 1 s
   "batch done confirmation" : Bool = PLC Batch_done_confirmation AT %M44.0, 1 s
   "Recipes_apporved" : Bool = PLC Rec_approved AT %M44.1, 1 s
   "Tank1_active" : Bool = PLC Tank1_active AT %M18.0, 1 s
   "valve A active" : Bool = PLC Valv_A_HMI AT %M18.2, 1 s
   "valve B active" : Bool = PLC Valv_B_HMI AT %M18.3, 1 s
   "valve C active" : Bool = PLC Valv_C_HMI AT %M18.4, 1 s
   "Drain valve active" : Bool = PLC Drain_valv_HMI AT %M18.6, 1 s
   "Agit_HMI" : Bool = PLC Agit_HMI AT %M18.5, 1 s
   "Alarm_active" : Bool = PLC Alarm_HMI AT %M18.1, 1 s

discrete alarms
   1: '', class Errors, trigger "Error_code" bit 0

text list "Alarm List": 999 'E-Stop Active'; 920 'Recipes not good'; 990 'Valve A Stuck Closed'; 980 'Valve B Stuck Closed'; 970 'Valve C stuck Closed'; 960 'Agitator Motor Didnt Start'; 950 'Drain Valve Stuck Open'; 940 'High level Over Flow'; 930 'Low Level Tank is empty'; 0 'No Alarm'

text list "Steps": 0 'Unit Ready'; 10 'Filling A'; 20 'Filling B'; 30 'FIlling C'; 40 'Agitating'; 50 'Draining'; 60 'waiting for Operator confirmation'; 999 'Unit Alarm'

recipe "Recipe": Recipe_element_A <- "Recipes_A", Recipe_element_B <- "Recipes_B", Recipe_element_C <- "Recipes_C"

screen "TAnk_1" 800x1280
   IOField "I/O field_1" at 601,1195 size 192x38; FormatPattern s999999999.999
      ProcessValue <- "Recipes_C"
   IOField "I/O field_2" at 601,1145 size 192x38; FormatPattern s999999999.999
      ProcessValue <- "Recipes_B"
   IOField "I/O field_3" at 601,1095 size 192x38; FormatPattern s999999999.999
      ProcessValue <- "Recipes_A"
   TextField "Text field_3" at 483,1203 size 85x27; Text 'Recipes C'
   TextField "Text field_4" at 483,1154 size 85x27; Text 'Recipes B'
   TextField "Text field_5" at 483,1105 size 85x27; Text 'Recipes A'
   Group "Group_2" at 483,1095 size 310x138
   Button "SB_NavigateHome_48x48" at 640,11 size 158x158; TextOff 'Text'; PictureOff "SB_NavigateHome_48x48_256c"
      on Click: ActivateScreen("home", 0)
   Switch "Pushbutton_Round_RN" at 25,1122 size 112x122; CaptionText 'Switch'; TextOff '0'; TextOn '1'; PictureOff "Pushbutton_Round_RN_Off_256c"; PictureOn "Pushbutton_Round_G_On_256c"
      ProcessValue <- "Start_Batch"
   Switch "Pushbutton_Round_RN_1" at 162,1122 size 112x122; CaptionText 'Switch'; TextOff '0'; TextOn '1'; PictureOff "Pushbutton_Round_RN_Off_256c"; PictureOn "Pushbutton_Round_G_On_256c"
      ProcessValue <- "Reset_HMI"
   Switch "Pushbutton_Round_RN_2" at 305,1122 size 112x122; CaptionText 'Switch'; TextOff '0'; TextOn '1'; PictureOn "Pushbutton_Round_N_On_mono"; PictureOff "Pushbutton_Round_RN_Off_256c"
      ProcessValue <- "batch done confirmation"
   TextField "Text field_1" at 25,1053 size 90x35; Text 'Start'
   TextField "Text field_2" at 162,1053 size 109x35; Text 'Reset'
   TextField "Text field_6" at 255,1055 size 182x35; Text 'Next Batch'
   Button "Button_4" at 10,29 size 235x48; TextOff 'Step TK1'
   Button "Button_7" at 318,29 size 235x48; TextOff 'Alarm 1'
      Appearance <- "Alarm_active"
   SymbolicIOField "Symbolic I/O field_2" at 10,92 size 234x32; TextOn '1'; TextOff '0'; TextList "Steps"
      ProcessValue <- "Status"
   SymbolicIOField "Symbolic I/O field_1" at 318,92 size 235x33; TextOn '1'; TextOff '0'; TextList "Alarm List"
      ProcessValue <- "Error_code"
   GraphicView "Graphic view_2" at 352,150 size 133x382; Picture "Graphic_17"
      Appearance <- "Agit_HMI"
   GraphicView "Graphic view_6" at 350,150 size 133x382; Picture "Graphic_21"
      Visibility <- "Agit_HMI"
   GraphicView "Graphic view_1" at 205,294 size 430x662; Picture "Graphic_16"
   Bar "Bar_1" at 304,360 size 68x582; MinimumValue 0; MaximumValue 500
      ProcessValue <- "level_value"
   Group "Group_3" at 614,418 size 83x96; Picture "Graphic_20"
   GraphicView "Graphic view_5" at 137,322 size 82x96; Picture "Graphic_20"
   GraphicView "Graphic view_7" at 134,322 size 82x96; Picture "Graphic_18"
      Visibility <- "valve A active"
   Group "Group" at 616,322 size 83x96; Picture "Graphic_20"
   GraphicView "Graphic view_10" at 134,846 size 82x96; Picture "Graphic_18"
      Visibility <- "Drain valve active"
   GraphicView "Graphic view_3" at 616,322 size 82x96; Picture "Graphic_20"
   GraphicView "Graphic view_4" at 617,322 size 82x96; Picture "Graphic_18"
      Visibility <- "valve B active"
   GraphicView "Graphic view_8" at 614,418 size 82x96; Picture "Graphic_20"
   GraphicView "Graphic view_9" at 615,418 size 82x96; Picture "Graphic_18"
      Visibility <- "valve C active"

screen "home" 800x1280
   Button "Button_1" at 20,46 size 235x48; TextOff 'TANK 1'
      on Press: ActivateScreen("TAnk_1", 0)
   Button "Button_2" at 287,46 size 235x48; TextOff 'TANK 2'
   Button "Button_3" at 547,46 size 235x48; TextOff 'TANK 3'
   IOField "I/O field_1" at 73,130 size 96x32; FormatPattern s999999999.999
      ProcessValue <- "level_value"
   IOField "I/O field_2" at 359,130 size 96x32; FormatPattern s999999999.999
      ProcessValue <- "level_value"
   IOField "I/O field_3" at 618,130 size 96x32; FormatPattern s999999999.999
      ProcessValue <- "level_value"
   Button "Button_4" at 20,217 size 235x48; TextOff 'Step TK1'
   Button "Button_5" at 287,217 size 235x48; TextOff 'Step TK2'
   Button "Button_6" at 547,217 size 235x48; TextOff 'Step TK3'
   IOField "I/O field_5" at 359,303 size 96x32; FormatPattern s99999
      ProcessValue <- "Status"
   IOField "I/O field_6" at 622,303 size 96x32; FormatPattern s99999
      ProcessValue <- "Status"
   Button "Button_7" at 20,382 size 235x48; TextOff 'Alarm 1'
      Appearance <- "Alarm_active"
      on Activate: function_fd9437ed(1, "Alarm_log_1")
   Button "Button_8" at 287,382 size 235x48; TextOff 'Alarm 2'
   Button "Button_9" at 547,382 size 235x48; TextOff 'Alarm 3'
   Button "Button_10" at 20,581 size 235x48; TextOff 'Config Tank1'; Authorization "User administration"
      on Press: ActivateScreen("Cnfig_tank_1", 0)
   Button "Button_11" at 287,581 size 235x48; TextOff 'Config Tank2'
   Button "Button_12" at 547,581 size 235x48; TextOff 'Config Tank3'
   Button "Button_13" at 20,700 size 235x48; TextOff 'REC Tank1'; Authorization "Supervisor"
      on Press: ActivateScreen("Receps", 0)
   Button "Button_14" at 287,700 size 235x48; TextOff 'REC Tank2'
   Button "Button_15" at 554,700 size 235x48; TextOff 'REC Tank3'
   Button "Button_16" at 616,1210 size 165x46; TextOff 'Login'
      on Press: ActivateScreen("LogIn", 0)
   Button "Button_17" at 434,1210 size 165x46; TextOff 'Alarm'
      on Press: ActivateScreen("Alarm_log", 0)
   SymbolicIOField "Symbolic I/O field_1" at 20,447 size 235x76; TextOff '0'; TextOn '1'; TextList "Alarm List"
      ProcessValue <- "Error_code"
   SymbolicIOField "Symbolic I/O field_2" at 11,303 size 257x32; TextOff '0'; TextOn '1'; TextList "Steps"
      ProcessValue <- "Status"

screen "Cnfig_tank_1" 800x1280
   Button "SB_NavigateHome_48x48" at 640,11 size 158x158; TextOff 'Text'; PictureOff "SB_NavigateHome_48x48_256c"
      on Click: ActivateScreen("home", 0)
   IOField "I/O field_1" at 528,303 size 240x34; FormatPattern s999999999.999
      ProcessValue <- "min_lvl"
   IOField "I/O field_2" at 528,253 size 240x34; FormatPattern s999999999.999
      ProcessValue <- "max _lvl"
   IOField "I/O field_3" at 528,353 size 240x34; FormatPattern s9999999999
      ProcessValue <- "Agitator_time_WD"
   IOField "I/O field_4" at 528,403 size 240x34; FormatPattern s9999999999
      ProcessValue <- "agitating_time"
   IOField "I/O field_5" at 528,453 size 240x34; FormatPattern s9999999999
      ProcessValue <- "filling_time_WD"
   IOField "I/O field_6" at 528,503 size 240x34; FormatPattern s9999999999
      ProcessValue <- "drain_time_WD"
   TextField "Text field_1" at 4,253 size 204x35; Text 'MAX_level'
   TextField "Text field_2" at 4,303 size 204x35; Text 'MIN_level'
   TextField "Text field_3" at 4,353 size 318x35; Text 'Agitator_timer_WD'
   TextField "Text field_4" at 4,403 size 318x35; Text 'Agitatiting_timr'
   TextField "Text field_5" at 4,453 size 318x35; Text 'Filling_timr_WD'
   TextField "Text field_6" at 4,503 size 318x35; Text 'Drain_Timr_Drain_'

screen "Receps" 800x1280
   IOField "I/O field_1" at 440,646 size 357x66; FormatPattern s999999999.999
      ProcessValue <- "Recipes_C"
   IOField "I/O field_2" at 438,422 size 357x66; FormatPattern s999999999.999
      ProcessValue <- "Recipes_B"
   IOField "I/O field_3" at 440,202 size 357x66; FormatPattern s999999999.999
      ProcessValue <- "Recipes_A"
   TextField "Text field_5" at 22,190 size 371x115; Text 'Recipes A'
   TextField "Text field_1" at 22,408 size 371x115; Text 'Recipes B'
   TextField "Text field_2" at 22,626 size 371x115; Text 'Recipes C'
   TextField "Text field_3" at 100,832 size 614x91; Text 'Recipes Approved'
   GraphicIOField "PlotLight_Round_G" at 266,992 size 246x216; PictureOn "PilotLight_Round_G_On_256c"; PictureOff "PilotLight_Round_G_Off_256c"
      ProcessValue <- "Recipes_apporved"
   Button "SB_NavigateHome_48x48" at 622,10 size 172x170; TextOff 'Text'; PictureOff "SB_NavigateHome_48x48_256c"
      on Click: ActivateScreen("home", 0)

screen "LogIn" 800x1280
   Button "Button_1" at 156,401 size 176x70; TextOff 'LogIn'
      on Press: function_a2a04561()
   Button "Button_2" at 428,401 size 190x71; TextOff 'LogOff'
      on Press: function_f23ef4c9()
   TextField "Text field_1" at 325,226 size 113x25; Text 'Current User'
   Button "SB_NavigateHome_48x48" at 622,10 size 172x170; TextOff 'Text'; PictureOff "SB_NavigateHome_48x48_256c"
      on Click: ActivateScreen("home", 0)

screen "Alarm_log" 800x1280
   Button "Button_2" at 547,1193 size 244x84; TextOff 'Home'
      on Press: ActivateScreen("home", 0)
   AlarmView "Alarm view_1" at 2,1 size 797x476; AlarmLog "Alarm_log_1"
*)